# B&R Automation Studio project MotorCylinder
Automation Studio 4.12.1

## Configuration Training

### Task classes (CPU.sw)
```
Cyclic#1 (cycle 10000 us):
  Main <- Main.prg
  Actuators <- Actuators.prg
```

### Hardware
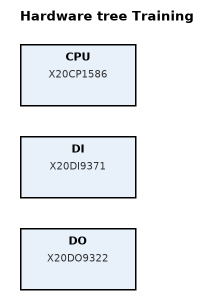
```
CPU : X20CP1586
  Cyclic1Duration = 10000
DI : X20DI9371
DO : X20DO9322
```

### IoMap.iom - CPU/IoMap.iom
```iecst
VAR_CONFIG
    StartButton AT %IX."DI".DigitalInput01;
    StopButton AT %IX."DI".DigitalInput02;
    DoorClosed AT %IX."DI".DigitalInput03;
    Motor1Running AT %IX."DI".DigitalInput04;
    Cylinder1Extended AT %IX."DI".DigitalInput05;
    Cylinder1Retracted AT %IX."DI".DigitalInput06;
    Motor1Cmd AT %QX."DO".DigitalOutput01;
    Cylinder1Extend AT %QX."DO".DigitalOutput02;
END_VAR
```

## Logical view

### Global.var
```iecst
VAR_GLOBAL
    StartButton : BOOL := FALSE;
    StopButton : BOOL := FALSE;
    DoorClosed : BOOL := TRUE;
    Motor1Cmd : BOOL := FALSE;
    Motor1Running : BOOL := FALSE;
    Cylinder1Extend : BOOL := FALSE;
    Cylinder1Extended : BOOL := FALSE;
    Cylinder1Retracted : BOOL := FALSE;
    Step : DINT := 0;
    CycleComplete : BOOL := FALSE;
END_VAR
```

### Program Logical/Actuators (IEC)

#### ActuatorsCyclic.st
```iecst
PROGRAM _CYCLIC
Motor1Cmd := (Step >= 1) AND (Step <= 3) AND DoorClosed;
Cylinder1Extend := (Step = 2) AND Motor1Running;
END_PROGRAM
```

### Program Logical/Main (IEC)

#### MainCyclic.st
```iecst
PROGRAM _CYCLIC
(* Training sequence. START is an explicit operator event. Feedback comes from the plant. *)
IF StopButton OR NOT DoorClosed THEN Step := 0; END_IF;
CASE Step OF
    0: IF StartButton AND DoorClosed AND Cylinder1Retracted THEN
           CycleComplete := FALSE; Step := 1;
       END_IF;
    1: IF Motor1Running THEN Step := 2; END_IF;
    2: IF Cylinder1Extended THEN Step := 3; END_IF;
    3: IF Cylinder1Retracted THEN CycleComplete := TRUE; Step := 4; END_IF;
END_CASE;
END_PROGRAM
```
